// TwinCAT 3 PLC project PLCStudent
// ProgramVersion: 3.1.4026.20
// libraries:
//   Tc2_Standard, * (Beckhoff Automation GmbH)
//   Tc2_System, * (Beckhoff Automation GmbH)
//   Tc3_Module, * (Beckhoff Automation GmbH)
// project tree:
//   / PlcTask.TcTTO
//   POUs/ BLINK.TcPOU, ControlFBD.TcPOU, MAIN.TcPOU
// (motion and I/O tree: see PLC project plcsim)
// real-time tasks:
//   TASK PlcTask: cycle T#30ms, priority 20, ADS port 350
// variable links:
//   PLCSim/PLCSim Instance <-> PLCStudent/PLCStudent Instance
//     PlcTask Inputs/MAIN.ixDrillDown <-> PlcTask Outputs/ControlFBD.qxDrillDown
//     PlcTask Inputs/MAIN.ixDrillUp <-> PlcTask Outputs/ControlFBD.qxDrillUp
//     PlcTask Inputs/MAIN.ixLampEmStopOk <-> PlcTask Outputs/ControlFBD.qxLampEmStopOk
//     PlcTask Inputs/MAIN.ixLampHomePos <-> PlcTask Outputs/ControlFBD.qxLampHomePos
//     PlcTask Inputs/MAIN.ixLampSafetyOk <-> PlcTask Outputs/ControlFBD.qxLampSafetyOk
//     PlcTask Inputs/MAIN.ixLampStarted <-> PlcTask Outputs/ControlFBD.qxLampStarted
//     PlcTask Inputs/MAIN.ixSliderAin <-> PlcTask Outputs/ControlFBD.qxSliderAin
//     PlcTask Inputs/MAIN.ixSliderAout <-> PlcTask Outputs/ControlFBD.qxSliderAout
//     PlcTask Inputs/MAIN.ixSliderBin <-> PlcTask Outputs/ControlFBD.qxSliderBin
//     PlcTask Inputs/MAIN.ixSliderBout <-> PlcTask Outputs/ControlFBD.qxSliderBout
//     PlcTask Outputs/MAIN.qxAuto <-> PlcTask Inputs/ControlFBD.ixAuto
//     PlcTask Outputs/MAIN.qxBtn1EmStopOk <-> PlcTask Inputs/ControlFBD.ixBtn1EmStopOk
//     PlcTask Outputs/MAIN.qxBtn2EmStopOk <-> PlcTask Inputs/ControlFBD.ixBtn2EmStopOk
//     PlcTask Outputs/MAIN.qxBtnAin <-> PlcTask Inputs/ControlFBD.ixBtnAin
//     PlcTask Outputs/MAIN.qxBtnAout <-> PlcTask Inputs/ControlFBD.ixBtnAout
//     PlcTask Outputs/MAIN.qxBtnBin <-> PlcTask Inputs/ControlFBD.ixBtnBin
//     PlcTask Outputs/MAIN.qxBtnBout <-> PlcTask Inputs/ControlFBD.ixBtnBout
//     PlcTask Outputs/MAIN.qxBtnDrillIn <-> PlcTask Inputs/ControlFBD.ixBtnDrillIn
//     PlcTask Outputs/MAIN.qxBtnDrillOut <-> PlcTask Inputs/ControlFBD.ixBtnDrillOut
//     PlcTask Outputs/MAIN.qxBtnReset <-> PlcTask Inputs/ControlFBD.ixBtnReset
//     PlcTask Outputs/MAIN.qxButtonStart <-> PlcTask Inputs/ControlFBD.ixButtonStart
//     PlcTask Outputs/MAIN.qxButtonStop <-> PlcTask Inputs/ControlFBD.ixButtonStop
//     PlcTask Outputs/MAIN.qxDrillDown <-> PlcTask Inputs/ControlFBD.ixDrillDown
//     PlcTask Outputs/MAIN.qxDrillUp <-> PlcTask Inputs/ControlFBD.ixDrillUp
//     PlcTask Outputs/MAIN.qxSafety1StopOk <-> PlcTask Inputs/ControlFBD.ixSafety1StopOk
//     PlcTask Outputs/MAIN.qxSafety2StopOk <-> PlcTask Inputs/ControlFBD.ixSafety2StopOk
//     PlcTask Outputs/MAIN.qxSliderAin <-> PlcTask Inputs/ControlFBD.ixSliderAin
//     PlcTask Outputs/MAIN.qxSliderAout <-> PlcTask Inputs/ControlFBD.ixSliderAout
//     PlcTask Outputs/MAIN.qxSliderBin <-> PlcTask Inputs/ControlFBD.ixSliderBin
//     PlcTask Outputs/MAIN.qxSliderBout <-> PlcTask Inputs/ControlFBD.ixSliderBout

CONFIGURATION PLCStudent
    RESOURCE PLC ON TwinCAT3
        TASK PlcTask(INTERVAL := T#30ms, PRIORITY := 20);
        PROGRAM MAIN WITH PlcTask : MAIN;
    END_RESOURCE
END_CONFIGURATION

// ---- POUs/MAIN.TcPOU
PROGRAM MAIN
VAR
END_VAR

ControlFBD();

END_PROGRAM

// ---- POUs/ControlFBD.TcPOU
PROGRAM ControlFBD
VAR
	qxLampStarted	AT %Q* : BOOL;
	qxSliderAout 	AT %Q* : BOOL; 
	qxSliderAin 	AT %Q* : BOOL; 
	qxSliderBout 	AT %Q* : BOOL; 
	qxSliderBin 	AT %Q* : BOOL; 
	qxDrillDown 	AT %Q* : BOOL;
	qxDrillUp		AT %Q* : BOOL;
	qxLampEmStopOk	AT %Q* : BOOL;
	qxLampSafetyOk  AT %Q* : BOOL;
	qxLampHomePos   AT %Q* : BOOL;
	
	
	mxManualRun : BOOL;
	mxEmergencyButtonPressed: BOOL;
	mxAuto : BOOL;
	mxAutoAIn : BOOL;
	mxAutoAOut : BOOL;
	mxAutoBIn : BOOL;
	mxAutoBOut : BOOL;
	mxAutoDrillDown: BOOL;
	mxAutoDrillUp: BOOL;
	
	mxSafetyOK : BOOL;
	mxManualOk : BOOL;
	mxCycleStopActivated : BOOL;
	mxBlink : BOOL;
	
	fbBlink : BLINK;

	
	
	ixButtonStart	AT %I* : BOOL;
	ixButtonStop	AT %I* : BOOL;
	ixSliderAout	AT %I* : BOOL;
	ixSliderAin		AT %I* : BOOL;
	ixSliderBout	AT %I* : BOOL;
	ixSliderBin		AT %I* : BOOL;
	ixDrillUp		AT %I* : BOOL;
	ixDrillDown		AT %I* : BOOL;

	ixAuto			AT %I* : BOOL;
	ixBtn1EmStopOk	AT %I* : BOOL;
	ixBtn2EmStopOk	AT %I* : BOOL;	
	ixSafety1StopOk	AT %I* : BOOL;
	ixSafety2StopOk	AT %I* : BOOL;	
	ixBtnReset		AT %I* : BOOL;
	ixBtnAout		AT %I* : BOOL;
	ixBtnAin		AT %I* : BOOL;
	ixBtnBout		AT %I* : BOOL;
	ixBtnBin		AT %I* : BOOL;
	ixBtnDrillOut	AT %I* : BOOL;
	ixBtnDrillIn	AT %I* : BOOL;

	mx: BOOL;
	mxStart: BOOL;
END_VAR

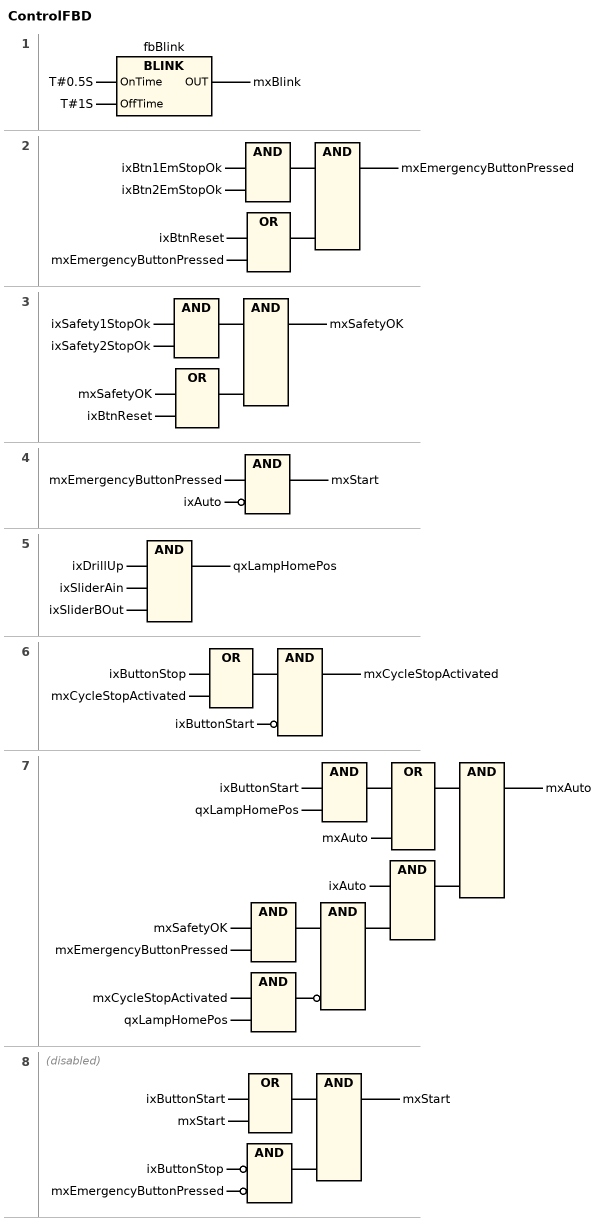
// NETWORK 1
fbBlink(OnTime := T#0.5S, OffTime := T#1S); // BLINK
mxBlink := fbBlink.OUT;

// NETWORK 2
mxEmergencyButtonPressed := (ixBtn1EmStopOk AND ixBtn2EmStopOk) AND (ixBtnReset OR mxEmergencyButtonPressed);

// NETWORK 3
mxSafetyOK := (ixSafety1StopOk AND ixSafety2StopOk) AND (mxSafetyOK OR ixBtnReset);

// NETWORK 4
mxStart := mxEmergencyButtonPressed AND NOT ixAuto;

// NETWORK 5
qxLampHomePos := ixDrillUp AND ixSliderAin AND ixSliderBOut;

// NETWORK 6
mxCycleStopActivated := (ixButtonStop OR mxCycleStopActivated) AND NOT ixButtonStart;

// NETWORK 7
mxAuto := (ixButtonStart AND qxLampHomePos OR mxAuto) AND (ixAuto AND ((mxSafetyOK AND mxEmergencyButtonPressed) AND NOT (mxCycleStopActivated AND qxLampHomePos)));

// NETWORK 8 (disabled)
// mxStart := (ixButtonStart OR mxStart) AND (NOT ixButtonStop AND NOT mxEmergencyButtonPressed);

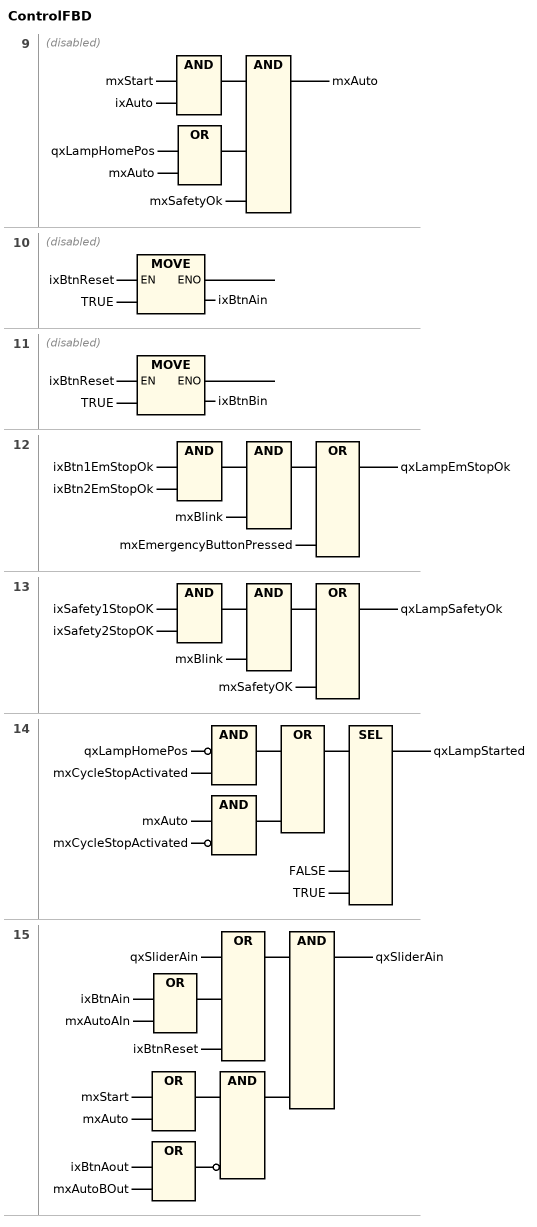
// NETWORK 9 (disabled)
// mxAuto := (mxStart AND ixAuto) AND (qxLampHomePos OR mxAuto) AND mxSafetyOk;

// NETWORK 10 (disabled)
// IF ixBtnReset THEN ixBtnAin := TRUE; END_IF

// NETWORK 11 (disabled)
// IF ixBtnReset THEN ixBtnBin := TRUE; END_IF

// NETWORK 12
qxLampEmStopOk := (ixBtn1EmStopOk AND ixBtn2EmStopOk) AND mxBlink OR mxEmergencyButtonPressed;

// NETWORK 13
qxLampSafetyOk := (ixSafety1StopOK AND ixSafety2StopOK) AND mxBlink OR mxSafetyOK;

// NETWORK 14
qxLampStarted := SEL(NOT qxLampHomePos AND mxCycleStopActivated OR mxAuto AND NOT mxCycleStopActivated, FALSE, TRUE);

// NETWORK 15
qxSliderAin := (qxSliderAin OR (ixBtnAin OR mxAutoAIn) OR ixBtnReset) AND ((mxStart OR mxAuto) AND NOT (ixBtnAout OR mxAutoBOut));

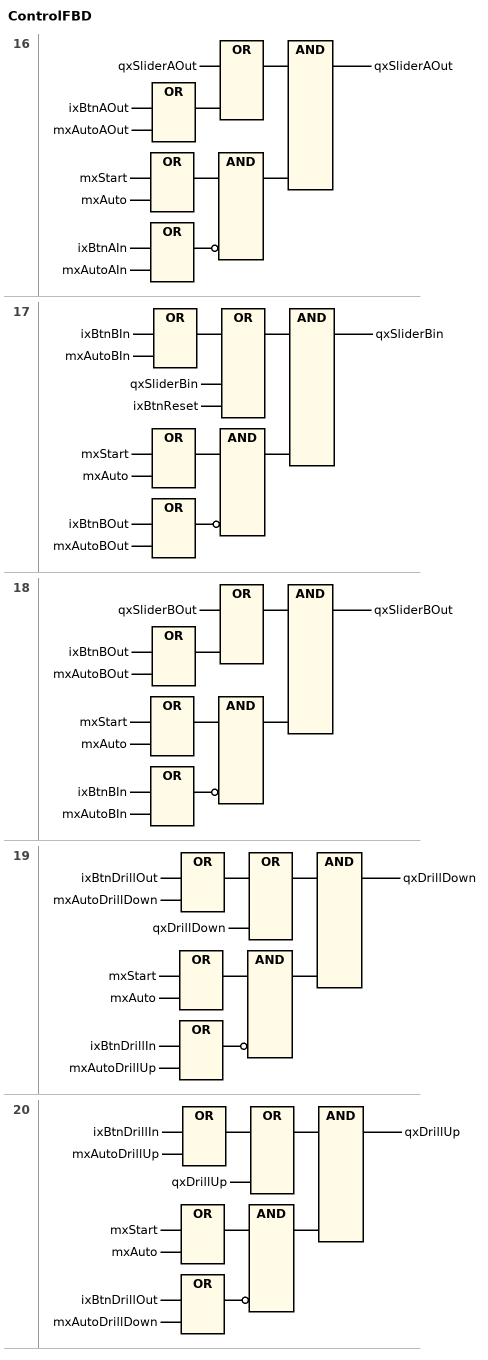
// NETWORK 16
qxSliderAOut := (qxSliderAOut OR (ixBtnAOut OR mxAutoAOut)) AND ((mxStart OR mxAuto) AND NOT (ixBtnAIn OR mxAutoAIn));

// NETWORK 17
qxSliderBin := ((ixBtnBIn OR mxAutoBIn) OR qxSliderBin OR ixBtnReset) AND ((mxStart OR mxAuto) AND NOT (ixBtnBOut OR mxAutoBOut));

// NETWORK 18
qxSliderBOut := (qxSliderBOut OR (ixBtnBOut OR mxAutoBOut)) AND ((mxStart OR mxAuto) AND NOT (ixBtnBIn OR mxAutoBIn));

// NETWORK 19
qxDrillDown := ((ixBtnDrillOut OR mxAutoDrillDown) OR qxDrillDown) AND ((mxStart OR mxAuto) AND NOT (ixBtnDrillIn OR mxAutoDrillUp));

// NETWORK 20
qxDrillUp := ((ixBtnDrillIn OR mxAutoDrillUp) OR qxDrillUp) AND ((mxStart OR mxAuto) AND NOT (ixBtnDrillOut OR mxAutoDrillDown));

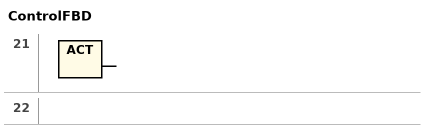
// NETWORK 21
ACT();

// NETWORK 22

ACTION ACT:
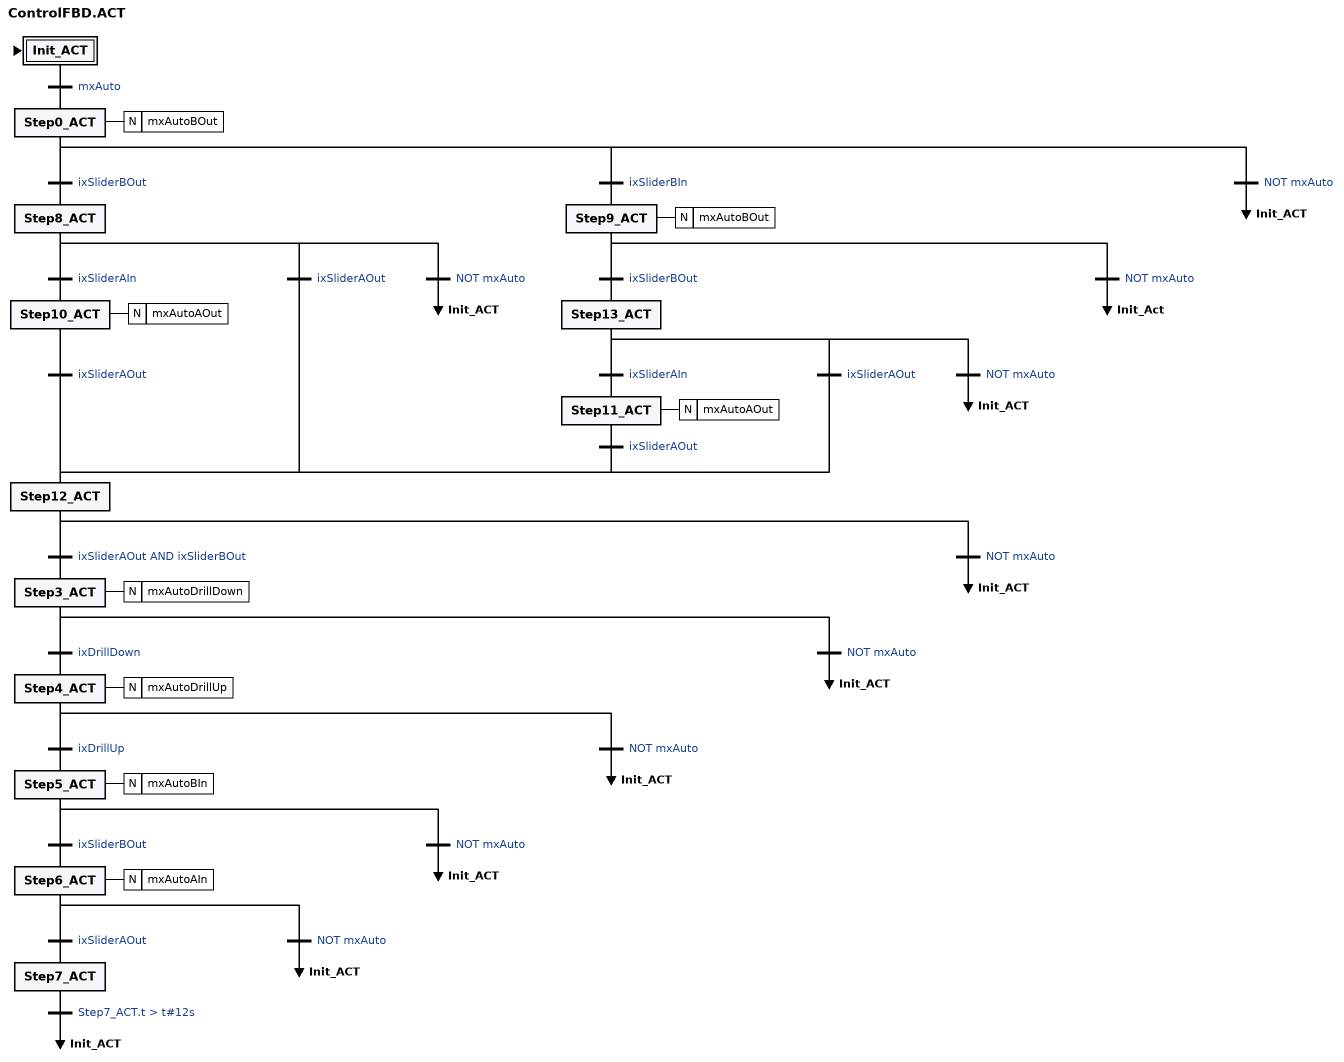
INITIAL_STEP Init_ACT:
END_STEP
TRANSITION FROM Init_ACT TO Step0_ACT
    := mxAuto;
END_TRANSITION
STEP Step0_ACT:
    mxAutoBOut(N);
END_STEP
TRANSITION FROM Step0_ACT TO Step8_ACT
    := ixSliderBOut;
END_TRANSITION
STEP Step8_ACT:
END_STEP
TRANSITION FROM Step8_ACT TO Step10_ACT
    := ixSliderAIn;
END_TRANSITION
STEP Step10_ACT:
    mxAutoAOut(N);
END_STEP
TRANSITION FROM Step10_ACT TO Step12_ACT
    := ixSliderAOut;
END_TRANSITION
TRANSITION FROM Step8_ACT TO Step12_ACT
    := ixSliderAOut;
END_TRANSITION
TRANSITION FROM Step8_ACT TO Init_ACT
    := NOT mxAuto;
END_TRANSITION
TRANSITION FROM Step0_ACT TO Step9_ACT
    := ixSliderBIn;
END_TRANSITION
STEP Step9_ACT:
    mxAutoBOut(N);
END_STEP
TRANSITION FROM Step9_ACT TO Step13_ACT
    := ixSliderBOut;
END_TRANSITION
TRANSITION FROM Step9_ACT TO Init_Act
    := NOT mxAuto;
END_TRANSITION
STEP Step13_ACT:
END_STEP
TRANSITION FROM Step13_ACT TO Step11_ACT
    := ixSliderAIn;
END_TRANSITION
STEP Step11_ACT:
    mxAutoAOut(N);
END_STEP
TRANSITION FROM Step11_ACT TO Step12_ACT
    := ixSliderAOut;
END_TRANSITION
TRANSITION FROM Step13_ACT TO Step12_ACT
    := ixSliderAOut;
END_TRANSITION
TRANSITION FROM Step13_ACT TO Init_ACT
    := NOT mxAuto;
END_TRANSITION
TRANSITION FROM Step0_ACT TO Init_ACT
    := NOT mxAuto;
END_TRANSITION
STEP Step12_ACT:
END_STEP
TRANSITION FROM Step12_ACT TO Step3_ACT
    := ixSliderAOut AND ixSliderBOut;
END_TRANSITION
TRANSITION FROM Step12_ACT TO Init_ACT
    := NOT mxAuto;
END_TRANSITION
STEP Step3_ACT:
    mxAutoDrillDown(N);
END_STEP
TRANSITION FROM Step3_ACT TO Step4_ACT
    := ixDrillDown;
END_TRANSITION
TRANSITION FROM Step3_ACT TO Init_ACT
    := NOT mxAuto;
END_TRANSITION
STEP Step4_ACT:
    mxAutoDrillUp(N);
END_STEP
TRANSITION FROM Step4_ACT TO Step5_ACT
    := ixDrillUp;
END_TRANSITION
TRANSITION FROM Step4_ACT TO Init_ACT
    := NOT mxAuto;
END_TRANSITION
STEP Step5_ACT:
    mxAutoBIn(N);
END_STEP
TRANSITION FROM Step5_ACT TO Step6_ACT
    := ixSliderBOut;
END_TRANSITION
TRANSITION FROM Step5_ACT TO Init_ACT
    := NOT mxAuto;
END_TRANSITION
STEP Step6_ACT:
    mxAutoAIn(N);
END_STEP
TRANSITION FROM Step6_ACT TO Step7_ACT
    := ixSliderAOut;
END_TRANSITION
TRANSITION FROM Step6_ACT TO Init_ACT
    := NOT mxAuto;
END_TRANSITION
STEP Step7_ACT:
END_STEP
TRANSITION FROM Step7_ACT TO Init_ACT
    := Step7_ACT.t > t#12s;
END_TRANSITION
// branch label Branch1_ACT
// branch label Branch3_ACT
// branch label Branch2_ACT
// branch label Branch0_ACT
// branch label Branch4_ACT
// branch label Branch5_ACT
// branch label Branch6_ACT
// branch label Branch7_ACT
// branch label Branch8_ACT
END_ACTION

ACTION Step14_ACT_exit:

END_ACTION

END_PROGRAM

// ---- POUs/BLINK.TcPOU
FUNCTION_BLOCK BLINK
VAR_INPUT
	OnTime : TIME;
	OffTime : TIME;
END_VAR
VAR_OUTPUT
	OUT : BOOL;
END_VAR
VAR
	fbTon : TON;
	fbOff : TON;
END_VAR

fbTon.PT := OnTime;
fbOff.PT := OffTime;

fbTon.IN := NOT fbOff.Q;
fbTon();

fboff.IN := fbOff.Q;
fbOff();

OUT := fbTon.Q;

END_FUNCTION_BLOCK
